// TIA Portal V21 export
DATA_BLOCK "Plant"   // DB41
{ S7_Optimized_Access := 'TRUE' }
// Motors supervised by PlantDiag.
   VAR
      pump : "Motor";
      fans : Array[0..1] of "Motor";
      count : Int;
   END_VAR
BEGIN
END_DATA_BLOCK
